Fanuc KAREL source: ko00063.KL

-- PROVISIONAL review KL for V1013-1; original PC SHA256 01f412e24a5f1c45422afa1b3778e92be0658b375a4697a5476adf6170f62880
-- Incomplete behavior may be omitted. Consult companion uncertainty JSON. Do not deploy.
PROGRAM KO00063
%NOLOCKGROUP
BEGIN
  -- UNRESOLVED_PC offsets 5-12; opcodes 9D,23
  -- UNRESOLVED_PC offsets 17-69; opcodes 27,27,49,7E,AD,27,49,7E,AD,22,31,7E,4A
  -- UNRESOLVED_PC offsets 74-78; opcodes 7F
END KO00063
